FUNCTION_BLOCK FB_GvlTest
VAR
	// Control
	nSeed : REFERENCE TO ULINT;

	// Private
	nLoopIndex1 : UDINT;
	nLoopIndex2 : UDINT;
END_VAR

// -----------------------------------------------------------------------
// Update variables — all fields are deterministic functions of seed
// -----------------------------------------------------------------------
GVL_Test.bBoolVar := (nSeed MOD 2 = 0);
GVL_Test.nSintVar := ULINT_TO_SINT(nSeed);
GVL_Test.nUsintVar := ULINT_TO_USINT(nSeed);
GVL_Test.nByteVar := ULINT_TO_BYTE(nSeed);
GVL_Test.nIntVar := ULINT_TO_INT(nSeed);
GVL_Test.nUintVar := ULINT_TO_UINT(nSeed);
GVL_Test.nWordVar := ULINT_TO_WORD(nSeed);
GVL_Test.nDintVar := ULINT_TO_DINT(nSeed);
GVL_Test.nUdintVar := ULINT_TO_UDINT(nSeed);
GVL_Test.nDwordVar := ULINT_TO_DWORD(nSeed);
GVL_Test.nLintVar := ULINT_TO_LINT(nSeed);
GVL_Test.nUlintVar := nSeed;
GVL_Test.nLwordVar := ULINT_TO_LWORD(nSeed);
GVL_Test.fRealVar := ULINT_TO_REAL(nSeed);
GVL_Test.fLrealVar := ULINT_TO_LREAL(nSeed);

// Date/time types — raw truncating casts, same bit pattern Go test will verify
GVL_Test.tTimeVar := ULINT_TO_TIME(nSeed);
GVL_Test.tdTimeOfDayVar := ULINT_TO_TOD(nSeed MOD 86400000);
GVL_Test.dDateVar := ULINT_TO_DATE(nSeed);
GVL_Test.dtDateTimeVar := ULINT_TO_DT(nSeed);
GVL_Test.tLTimeVar := ULINT_TO_LTIME(nSeed);
GVL_Test.tdLTimeOfDayVar  := ULINT_TO_LTOD(nSeed MOD 86400000000000);
GVL_Test.dLDateVar := ULINT_TO_LDATE(nSeed);
GVL_Test.dtLDateTimeVar := ULINT_TO_LDT(nSeed);
GVL_Test.sStringVar := CONCAT('S=', ULINT_TO_STRING(nSeed));

// -----------------------------------------------------------------------
// Update test struct — all fields are deterministic functions of seed
// -----------------------------------------------------------------------
GVL_Test.stStructVar.nSeed := ULINT_TO_UDINT(nSeed);
GVL_Test.stStructVar.bBoolVar := GVL_Test.bBoolVar;
GVL_Test.stStructVar.nSintVar := GVL_Test.nSintVar;
GVL_Test.stStructVar.nUsintVar := GVL_Test.nUsintVar;
GVL_Test.stStructVar.nByteVar := GVL_Test.nByteVar;
GVL_Test.stStructVar.nIntVar := GVL_Test.nIntVar;
GVL_Test.stStructVar.nUintVar := GVL_Test.nUintVar;
GVL_Test.stStructVar.nWordVar := GVL_Test.nWordVar;
GVL_Test.stStructVar.nDintVar := GVL_Test.nDintVar;
GVL_Test.stStructVar.nUdintVar := GVL_Test.nUdintVar;
GVL_Test.stStructVar.nDwordVar := GVL_Test.nDwordVar;
GVL_Test.stStructVar.nLintVar := GVL_Test.nLintVar;
GVL_Test.stStructVar.nUlintVar := GVL_Test.nUlintVar;
GVL_Test.stStructVar.nLwordVar := GVL_Test.nLwordVar;
GVL_Test.stStructVar.fRealVar := GVL_Test.fRealVar;
GVL_Test.stStructVar.fLrealVar := GVL_Test.fLrealVar;
GVL_Test.stStructVar.tTimeVar := GVL_Test.tTimeVar;
GVL_Test.stStructVar.tdTimeOfDayVar := GVL_Test.tdTimeOfDayVar;
GVL_Test.stStructVar.dDateVar := GVL_Test.dDateVar;
GVL_Test.stStructVar.dtDateTimeVar := GVL_Test.dtDateTimeVar;
GVL_Test.stStructVar.tLTimeVar := GVL_Test.tLTimeVar;
GVL_Test.stStructVar.tdLTimeOfDayVar := GVL_Test.tdLTimeOfDayVar;
GVL_Test.stStructVar.dLDateVar := GVL_Test.dLDateVar;
GVL_Test.stStructVar.dtLDateTimeVar := GVL_Test.dtLDateTimeVar;
GVL_Test.stStructVar.sStringVar := GVL_Test.sStringVar;

// -----------------------------------------------------------------------
// Update 1-D arrays: element[i] = UDINT_TO_x(seed + i)
// -----------------------------------------------------------------------
FOR nLoopIndex1 := 0 TO 9 DO
	GVL_Test.aIntArray[nLoopIndex1] := ULINT_TO_INT(nSeed + nLoopIndex1);
	GVL_Test.aDintArray[nLoopIndex1] := ULINT_TO_DINT(nSeed + nLoopIndex1);
END_FOR

// -----------------------------------------------------------------------
// Update 2-D array: element[i,j] = UDINT_TO_INT(seed + i*3 + j)
// -----------------------------------------------------------------------
FOR nLoopIndex1 := 0 TO 2 DO
	FOR nLoopIndex2 := 0 TO 2 DO
		GVL_Test.aIntArray2d[nLoopIndex1, nLoopIndex2] := ULINT_TO_INT(nSeed + nLoopIndex1 * 3 + nLoopIndex2);
	END_FOR
END_FOR

//FB_Init is always available implicitly and it is used primarily for initialization.
//The return value is not evaluated. For a specific influence, you can also declare the
//methods explicitly and provide additional code there with the standard initialization
//code. You can evaluate the return value.
METHOD FB_Init: BOOL
VAR_INPUT
    bInitRetains : BOOL; // TRUE: the retain variables are initialized (reset warm / reset cold)
    bInCopyCode : BOOL;  // TRUE: the instance will be copied to the copy code afterward (online change)
	nSeed : REFERENCE TO ULINT;
END_VAR
THIS^.nSeed REF= nSeed;
END_METHOD

END_FUNCTION_BLOCK

(* stored: Version 1.1.0.1, ProductVersion 3.1.4026.19
   POU FB_GvlTest: Id {e64978a6-7b94-4bc8-a366-3a9a51ec0fb5}, SpecialFunc None
   Method FB_Init: Id {8b66484e-bb4e-4270-b0d2-b32177d32d63} *)
